(* IEC 61131-3 sources: llm-plc-st-eval/data/processed_definitivo/claude-sonnet-4-6/C8/zero_shot, 3 files *)

(* ---- ejec_1.st ---- *)
FUNCTION_BLOCK FB_Valvula
VAR_INPUT
    nivelAlto : BOOL; (* Señal de nivel alto *)
END_VAR

VAR_OUTPUT
    valvula : BOOL; (* Salida hacia la válvula *)
END_VAR

VAR
    T1 : TON; (* Temporizador a la conexión, retardo a la activación *)
END_VAR

(* -------------------------------------------------------
   Rama 1: nivelAlto activa el temporizador T1 (TON, PT=5s)
   Rama 2: cuando T1.Q=TRUE se activa la salida valvula
   ------------------------------------------------------- *)

(* Rama 1: equivalente al contacto NA nivelAlto -> TON T1 *)
T1(IN := nivelAlto, PT := T#5S);

(* Rama 2: equivalente al contacto NA T1.Q -> bobina valvula *)
valvula := T1.Q;
END_FUNCTION_BLOCK

(* ---- ejec_2.st ---- *)
FUNCTION_BLOCK FB_Valvula
VAR_INPUT
    nivelAlto : BOOL; (* Sensor de nivel alto *)
END_VAR

VAR_OUTPUT
    valvula : BOOL; (* Bobina de la válvula *)
END_VAR

VAR
    T1 : TON; (* Temporizador a la conexión, retardo a la conexión *)
END_VAR

(* -------------------------------------------------------
   Rama 1: nivelAlto activa el temporizador T1 (TON, PT = 5 s)
   Rama 2: T1.Q activa la bobina valvula
   ------------------------------------------------------- *)

(* Rama 1 - Temporizador TON *)
T1(IN := nivelAlto, PT := T#5S);

(* Rama 2 - Bobina valvula *)
valvula := T1.Q;
END_FUNCTION_BLOCK

(* ---- ejec_3.st ---- *)
FUNCTION_BLOCK FB_Valvula
VAR_INPUT
    nivelAlto : BOOL; (* Señal de nivel alto *)
END_VAR

VAR_OUTPUT
    valvula : BOOL; (* Salida hacia la válvula *)
END_VAR

VAR
    T1 : TON; (* Temporizador a la conexión, 5 segundos *)
END_VAR

(* Rama 1: nivelAlto activa el temporizador T1 con PT = 5 s *)
T1(IN := nivelAlto, PT := T#5S);

(* Rama 2: cuando T1 expira (Q = TRUE), se activa la válvula *)
valvula := T1.Q;
